(* IEC 61131-3 sources: PLC-Static-Analysis/modules/plc-rules/src/test/resources/PLCA-L010, 2 files *)

(* ---- compliant.st ---- *)
FUNCTION F_Next : INT
F_Next := 1;
END_FUNCTION

PROGRAM P_L010ok
VAR
    n : INT;
    m : INT;
    r : REAL;
    b : BOOL;
    c : BOOL;
    q : BOOL;
END_VAR
IF n > 10 AND n < 50 THEN
    q := TRUE;
END_IF
q := F_Next() > 10 AND F_Next() > 5;
q := b AND c;
q := (b OR c) AND NOT b;
END_PROGRAM

(* ---- noncompliant.st ---- *)
PROGRAM P_L010
VAR
    n : INT;
    m : INT;
    r : REAL;
    b : BOOL;
    c : BOOL;
    q : BOOL;
END_VAR
IF n > 10 AND n > 5 THEN // PLCA-L010
    q := TRUE;
END_IF
q := n > 10 OR n > 5; // PLCA-L010
q := b AND c AND b; // PLCA-L010
q := (b OR c) AND b; // PLCA-L010
END_PROGRAM
